Fanuc KAREL source: KT00474.KL

PROGRAM KT00474
%NOLOCKGROUP
VAR
  P1: POSITION
  P2: POSITION
  OUT: POSITION
BEGIN
  OUT = P1 : P2
END KT00474
